Fanuc KAREL source: KC00024.KL

PROGRAM KC00024
%NOLOCKGROUP
VAR
  I: INTEGER
  J: INTEGER
  K: INTEGER
  R: REAL
  B: BOOLEAN
  S: STRING[80]
  T: STRING[80]
  P: PATH
  Q: PATH
  AI: ARRAY[8] OF INTEGER
  AB: ARRAY[244] OF BYTE
BEGIN
  S = ''
  T = 'I'
  DAQ_REGPIPE(1,1,10,S,T,S,1,J)
END KC00024
